FUNCTION F_atan2 : REAL
VAR_INPUT
	rX	:	REAL;
	rY	:	REAL;
END_VAR
VAR
END_VAR

// CALCOLO L'ANGOLO CONOSCENDO COORDINATE X E Y
IF rX > 0 THEN
	F_atan2	:=	ATAN(rY / rX);
ELSIF rX = 0 AND rY > 0 THEN
	F_atan2	:=	LREAL_TO_REAL(CONSTANTS.PI / 2);
ELSIF rX = 0 AND rY < 0 THEN
	F_atan2	:=	- LREAL_TO_REAL(CONSTANTS.PI / 2);
ELSIF rX < 0 AND rY >= 0 THEN
	F_atan2	:=	LREAL_TO_REAL(ATAN(rY / rX) + CONSTANTS.PI);
ELSIF rX < 0 AND rY < 0 THEN
	F_atan2	:=	LREAL_TO_REAL(ATAN(rY / rX) - CONSTANTS.PI);
END_IF

END_FUNCTION

(* stored: Version 1.1.0.1, ProductVersion 3.1.4024.9
   POU F_atan2: Id {b2c16367-73dd-4a68-96c2-1c66916166e8}, SpecialFunc None *)
